Fanuc KAREL source: KT00845.KL

PROGRAM KT00845
%NOLOCKGROUP
VAR
  I1: INTEGER
  I2: INTEGER
  OUT: REAL
BEGIN
  I1 = 2
  I2 = 3
  I1 = 2
  I2 = 3
  OUT = TAN(I1)
END KT00845
